Staubli VAL3: LibTorque.dtx

public bool bDisable[4]
  [0] = true
  [1] = true
  [2] = true
  [3] = true
bool bLock
bool bSix_Axis
mdesc mNomSpeed
num nCurrentMaxForce
public num nMaxJntForce[4]
  [0] = 1000000
  [1] = 1000000
  [2] = 21.1
  [3] = 65
num nMaxJntGet
string sArm4List[9]
  [0] = "tp_80"
  [1] = "ts2_100"
  [2] = "ts2_40"
  [3] = "ts2_60"
  [4] = "ts2_80"
  [5] = "ts_20"
  [6] = "ts_40"
  [7] = "ts_60"
  [8] = "ts_80"
string sArm6List[16]
  [0] = "rx_160"
  [1] = "tx2_140"
  [2] = "tx2_160"
  [3] = "tx2_160l"
  [4] = "tx2_200"
  [5] = "tx2_200l"
  [6] = "tx2_40"
  [7] = "tx2_60"
  [8] = "tx2_60l"
  [9] = "tx2_90"
  [10] = "tx2_90l"
  [11] = "tx2_90xl"
  [12] = "tx_200"
  [13] = "tx_40"
  [14] = "tx_60"
  [15] = "tx_90"
string sArmDetail = "ts2_40"
string sArmType = "4_Axis"
public string sBtnUnLock = "保存"
string sPassword = "staubli2025"
